Fanuc KAREL source: kt00402.KL

-- PROVISIONAL review KL for V940-1; original PC SHA256 d49141ffcb7a7448f6ac943b5ee10eb0652a68d817ce3b40d2dc5f9c21ce0d3d
-- Incomplete behavior may be omitted. Consult companion uncertainty JSON. Do not deploy.
PROGRAM KT00402
%NOLOCKGROUP
VAR
  I1 : INTEGER
  R2 : REAL
  OUT : BOOLEAN
BEGIN
  -- V9_ZERO_TABLE_METADATA_HINT layout=0001; no indexed target words; source/name/runtime held
  -- UNRESOLVED_PC offsets 5-16; opcodes 2E,23
  -- UNRESOLVED_PC offsets 21-32; opcodes 2E,23
  -- UNRESOLVED_PC offsets 37-59; opcodes 21,21,29,64,29,71,23
  -- UNRESOLVED_PC offsets 64-68; opcodes 7F
END KT00402
